(* IEC 61131-3 sources: plc-vscode/tests/st/test-ready/rusty/tests/lit/multi/variable_length_array_size, 3 files *)

(* ---- function.st ---- *)
FUNCTION function_1 : INT
VAR_INPUT
    x3 : ARRAY [*] OF INT;
END_VAR
VAR_OUTPUT
    x4 : ARRAY [*,*] OF INT;
END_VAR
VAR_IN_OUT
    x5 : ARRAY [*,*] OF INT;
END_VAR
VAR
END_VAR
    printf('Test$N');
    function_1 := 0;
END_FUNCTION

(* ---- main.st ---- *)
FUNCTION main
    VAR
        fb1: function_block_1;
        arr: ARRAY[0..14, -2..1] OF INT;
        arr2: ARRAY[0..14] OF INT;
        arr3: ARRAY[0..14, -2..1] OF INT;
        arr4: ARRAY[0..14, -2..1] OF INT;
    END_VAR

    fb1(arr);
    function_1(arr2, arr3, arr4);
END_FUNCTION

(* ---- function_block.st ---- *)
FUNCTION_BLOCK function_block_1
VAR_INPUT
END_VAR
VAR_OUTPUT
END_VAR
VAR_IN_OUT
    x1 : ARRAY [*,*] OF INT;
END_VAR
VAR
END_VAR
END_FUNCTION_BLOCK
